FUNCTION_BLOCK FB_EL3351ChannelDiagnosis_1
VAR_INPUT
	stBridgeState					:ST_EL3351ChannelState;				(* AI bridge state *)
	stSupplyState					:ST_EL3351ChannelState;				(* AI supply state *)
END_VAR
VAR_OUTPUT
	bBridgeChannelOK			:BOOL;
	bSupplyChannelOK			:BOOL;
END_VAR
VAR

END_VAR


(* General Channel Status *)
IF stBridgeState.bUnderrange= 0
    AND stBridgeState.bOverrangerange= 0
    AND stBridgeState.bError= 0
    AND stBridgeState.bState= 0
THEN
	bBridgeChannelOK:= TRUE;
ELSE
	bBridgeChannelOK:= FALSE;
END_IF

IF stSupplyState.bUnderrange= 0
     AND stSupplyState.bOverrangerange= 0
     AND stSupplyState.bError= 0
     AND stSupplyState.bState= 0
THEN
	bSupplyChannelOK:= TRUE;
ELSE
	bSupplyChannelOK:= FALSE;
END_IF

END_FUNCTION_BLOCK

(* stored: Version 1.1.0.1, ProductVersion 3.1.4024.15
   POU FB_EL3351ChannelDiagnosis_1: Id {80e89fa4-6758-463c-9f9a-415d530ddf47}, SpecialFunc None *)
